(* IEC 61131-3 sources: plc-iiot-stack/src/POUs/Iiot/F_IiotClockValid, 1 file *)

(* ---- F_IiotClockValid.decl.st ---- *)
// Назначение: время ПЛК в диапазоне ts схемы (2020-01-01 .. 2100-01-01 UTC): без этого сообщения
//             были бы вне схемы, и обмен не начинается.
// Автор:      kr0nsch
// Версия:     0.1.0
// Документ:   docs/plc_mqtt.md, раздел «Связь и состояние узла»
FUNCTION F_IiotClockValid : BOOL
VAR_INPUT
    uliTs_ms : ULINT;   // мс от 1970-01-01 UTC
END_VAR
